{attribute 'linkalways'}
{attribute 'no_explicit_call' := 'Use the methods of this class'}
{attribute 'enable_dynamic_creation'}
FUNCTION_BLOCK Lidar_Watchdog IMPLEMENTS I_Lidar
VAR
	timeoutError : HardwareError := (isActive := TRUE, id := Constants.LIDAR_TIMEOUT_ERROR_ID, text := 'Ingen LIDAR-skann innenfor fristen');
	inner : I_Lidar;
	timeoutTimer : TON;
	isTimedOut : BOOL;
END_VAR

METHOD Wrap
VAR_INPUT
	lidar : I_Lidar;
END_VAR
inner := lidar;
END_METHOD

METHOD Execute
IF inner = 0 THEN
	RETURN;
END_IF
timeoutTimer(IN := inner.IsRunning, PT := Constants.LIDAR_TIMEOUT_IN_MS);
IF timeoutTimer.Q THEN
	isTimedOut := TRUE;
END_IF
END_METHOD

METHOD Start
IF inner <> 0 THEN
	inner.Start();
END_IF
timeoutTimer(IN := FALSE);
isTimedOut := FALSE;
END_METHOD

METHOD Stop
IF inner <> 0 THEN
	inner.Stop();
END_IF
timeoutTimer(IN := FALSE);
isTimedOut := FALSE;
END_METHOD

METHOD TryGetScan : BOOL
VAR_INPUT
	scan : REFERENCE TO LaserScan;
END_VAR
IF inner = 0 OR_ELSE NOT inner.TryGetScan(scan) THEN
	RETURN;
END_IF
timeoutTimer(IN := FALSE);
isTimedOut := FALSE;
TryGetScan := TRUE;
END_METHOD

PROPERTY IsRunning : BOOL
GET
IsRunning := inner <> 0 AND_THEN inner.IsRunning;
END_GET
END_PROPERTY

PROPERTY Error : HardwareError
GET
IF isTimedOut THEN
	Error := timeoutError;
ELSIF inner <> 0 THEN
	Error := inner.Error;
END_IF
END_GET
END_PROPERTY

END_FUNCTION_BLOCK

(* stored: Version 1.1.0.1, ProductVersion 3.1.4026.12
   POU Lidar_Watchdog: Id {11055b29-6e9e-5314-983d-7ebae39fc2b9}, SpecialFunc None
   Method Wrap: Id {b8d46fca-05a4-56f2-8cb0-d35ef837e6f7}
   Method Execute: Id {1f8caded-dcfd-5177-afdb-eccd18e79341}
   Method Start: Id {8882ed4d-3a47-5d6e-b86e-9f8693655116}
   Method Stop: Id {f2da4acb-3f55-5b16-be8a-4d1ea57efd3c}
   Method TryGetScan: Id {fff34688-a6e0-5382-9d37-5023f230c7ab}
   Property IsRunning: Id {2c63264d-d2c8-587c-9556-76232fb1faa0}
   Get Get: Id {9c1f7fce-392c-5756-92e0-e337b7ba4617}
   Property Error: Id {5092db6b-38c6-5d81-9352-19c8af0a3350}
   Get Get: Id {ed4fe3fb-6d61-5641-9107-5cea4f8caf09} *)
